(* Logix 5000 project; controller RV_2AJ 1769-L16ER-BB1B rev 36.11; software revision 36.00 *)

TASK MainTask (continuous, watchdog 500 ms) : MainProgram

MODULES
   Local : 1769-L16ER-BB1B (PointIO 0, rev 36.11)
      Input_1_Sink : 1734-IB8 (PointIO 5, rev 3.1, Input RPI 20 ms)
           Local:5:I.Data.0   // Slide_Sensor
           Local:5:I.Data.1   // Hand_Sensor
           Local:5:I.Data.2   // Block_Sensor
      Input_2_Source : 1734-IV8 (PointIO 6, rev 3.1, Input RPI 20 ms)
      Discrete_IO : Embedded (PointIO 1, rev 36.11, Output RPI 20 ms)
           Local:1:I.Data.0   // Robot_Running
           Local:1:I.Data.1   // Robot_Servo_On
           Local:1:I.Data.10   // Open
           Local:1:I.Data.11   // Open
           Local:1:I.Data.12   // Open
           Local:1:I.Data.13   // Open
           Local:1:I.Data.14   // Open
           Local:1:I.Data.15   // Open
           Local:1:I.Data.2   // Robot_Error
           Local:1:I.Data.3   // Robot_Operation_Rights
           Local:1:I.Data.4   // Open
           Local:1:I.Data.5   // Open
           Local:1:I.Data.6   // Open
           Local:1:I.Data.7   // Open
           Local:1:I.Data.8   // Open
           Local:1:I.Data.9   // Open
           Local:1:O.Data.0   // Robot_Stop(All Slot)
           Local:1:O.Data.1   // Robot_ Servo_Off
           Local:1:O.Data.10   // Block_Sensor
           Local:1:O.Data.11   // Open
           Local:1:O.Data.12   // Open
           Local:1:O.Data.13   // Open
           Local:1:O.Data.14   // Open
           Local:1:O.Data.15   // Open
           Local:1:O.Data.2   // Robot_ Error_Reset
           Local:1:O.Data.3   // Robot_Start
           Local:1:O.Data.4   // Robot_ Servo_On
           Local:1:O.Data.5   // Robot_Opertion_Rights
           Local:1:O.Data.6   // Open
           Local:1:O.Data.7   // Open
           Local:1:O.Data.8   // Slide_Sensor
           Local:1:O.Data.9   // Hand_Sensor
      Out_2 : 1734-OW4 (PointIO 3, rev 3.1, Output RPI 20 ms)
      Out_3 : 1734-OW4 (PointIO 4, rev 3.1, Output RPI 20 ms)
      Out_1 : 1734-OW4 (PointIO 2, rev 3.1, Output RPI 20 ms)
END_MODULES

VAR_GLOBAL   (* controller tags *)
   T4_0 : TIMER := (PRE := 35000);   // Test_Timer
END_VAR

PROGRAM MainProgram   (* main routine MainRoutine *)
VAR
   Robot_Finished : BOOL;
   Trigger_Wave : BOOL;
END_VAR

ROUTINE MainRoutine   (* ladder *)
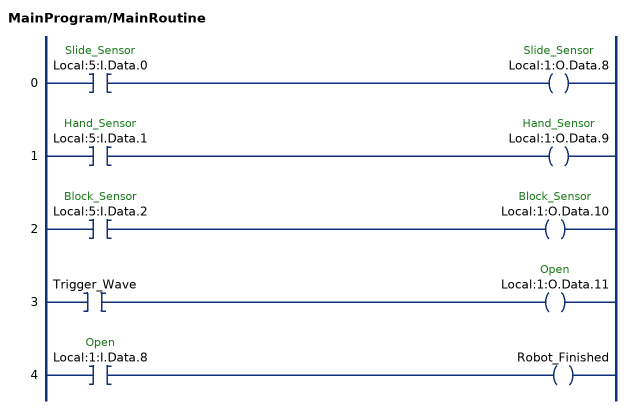
   0: XIC(Local:5:I.Data.0)OTE(Local:1:O.Data.8);
   1: XIC(Local:5:I.Data.1)OTE(Local:1:O.Data.9);
   2: XIC(Local:5:I.Data.2)OTE(Local:1:O.Data.10);
   3: XIC(Trigger_Wave)OTE(Local:1:O.Data.11);
   4: XIC(Local:1:I.Data.8)OTE(Robot_Finished);
END_ROUTINE
END_PROGRAM
